// TIA Portal project "Dual_Pump_Pressure_Control" (V20)

(* hardware
DEVICE "S7-1500/ET200MP station_1"  S7-1500 station
   slot 0: "Rail_0"  Rack  6ES7 590-1***0-0AA0
   slot 1: "PLC_PumpStation"  CPU 1511-1 PN  6ES7 511-1AL03-0AB0  V4.0
      slot 3: "CPU display_1"  6ES7591-1AA00-0AA0
      slot 32768: "PROFINET interface_1"  X1
         slot 32769: "Port_1"  X1 P1
         slot 32770: "Port_2"  X1 P2
      slot 34817: "Virtual CP interface port_1"  Virtual CP interface port  Virtual CP interface port FW V4.0
DEVICE "HMI_PumpStation"  TP1500 Comfort
   slot 0: "HMI_PumpStation"  TP1500 Comfort  6AV2 124-0QC02-0AX0  17.0.0.0
   slot 1: "HMI_RT_1"  TP1500 Comfort  6AV2 124-0QC02-0AX0  17.0.0.0
   slot 5: "HMI_PumpStation.IE_CP_1"  PROFINET Interface  17.0.0.0
      slot 1: "PROFINET Interface_1"  PROFINET Interface
         slot 1: "Port_1"  Port
         slot 2: "Port_2"  Port
   slot 6: "HMI_PumpStation.IE_CP_2"  PROFINET Interface  17.0.0.0
      slot 1: "PROFINET Interface_GBit"  PROFINET Interface
         slot 1: "Port_1"  Port
   slot 7: "HMI_PumpStation.MPI/DP_CP_1"  MPI/DP Interface  17.0.0.0
DEVICE "SCADA_PumpStation"  SIMATIC PC station
   slot 0: "SIMATIC PC station"  Rail  SIMATIC PC-Station  V1.0
      slot 125: "Stationmanager"  Station_Manager  V6.0.4
   slot 1: "HMI_RT_2"  WinCC Unified PC RT  6AV2 155-xxxxx-xxxx  20.0.0.0
   slot 2: "IE general_1"  IE General  IE_CP  V8.2.0
      slot 1: "PROFINET interface"  IEGeneral.Interface.8.2.0
*)

// ===== PLC "PLC_PumpStation"  CPU 1511-1 PN =====

DATA_BLOCK "DB_Sim"   // DB1
{ S7_Optimized_Access := 'TRUE' }
VERSION : 0.1
   VAR
      Water_Level_OK : Bool := true;
      P1_InjectFault : Bool;
      P2_InjectFault : Bool;
   END_VAR
BEGIN
END_DATA_BLOCK

DATA_BLOCK "DB_IO"   // DB2
{ S7_Optimized_Access := 'TRUE' }
VERSION : 0.1
   VAR
      P1_RunCmd : Bool;
      P1_Speed_SP : Real := 0.0;
      P1_Ready : Bool;
      P1_RunningFB : Bool;
      P1_StoppedFB : Bool;
      P1_Fault : Bool;
      P2_RunCmd : Bool;
      P2_Speed_SP : Real;
      P2_Ready : Bool;
      P2_RunningFB : Bool;
      P2_StoppedFB : Bool;
      P2_Fault : Bool;
      P1_Status : Int;
      P2_Status : Int;
      AnyPumpRunning : Bool;
      Pressure_PV : Real;
      PID_Output : Real;
      PID_Enable : Bool;
      PID_Reset : Bool;
      PID_Mode : Int := 3;
   END_VAR
BEGIN
END_DATA_BLOCK

DATA_BLOCK "DB_VFD_Sim_P1"   // DB3
{ S7_Optimized_Access := 'TRUE' }
VERSION : 0.1
// stored: InstanceOfName FB_VFD_Sim
"FB_VFD_Sim"
BEGIN
END_DATA_BLOCK

DATA_BLOCK "DB_VFD_Sim_P2"   // DB4
{ S7_Optimized_Access := 'TRUE' }
VERSION : 0.1
// stored: InstanceOfName FB_VFD_Sim
"FB_VFD_Sim"
BEGIN
END_DATA_BLOCK

DATA_BLOCK "DB_HMI"   // DB5
{ S7_Optimized_Access := 'TRUE' }
VERSION : 0.1
   VAR
      Cmd_AutoMode : Bool;
      Cmd_Start : Bool;
      Cmd_Stop : Bool;
      Cmd_ManualPump : USInt := 1;
      Cmd_ManualSpeed_SP : Real := 50.0;
      Cmd_SystemReset : Bool;
      Pressure_SP : Real := 6.0;
   END_VAR
BEGIN
END_DATA_BLOCK

DATA_BLOCK "DB_PumpStation"   // DB6
{ S7_Optimized_Access := 'TRUE' }
VERSION : 0.1
// stored: InstanceOfName FB_PumpStation
"FB_PumpStation"
BEGIN
END_DATA_BLOCK

DATA_BLOCK "DB_Process_Sim"   // DB7
{ S7_Optimized_Access := 'TRUE' }
VERSION : 0.1
// stored: InstanceOfName FB_Process_Sim
"FB_Process_Sim"
BEGIN
END_DATA_BLOCK

DATA_BLOCK "DB_Alarms"   // DB9
{ S7_Optimized_Access := 'TRUE' }
VERSION : 0.1
   VAR
      AlarmWord : Word;
   END_VAR
BEGIN
END_DATA_BLOCK

FUNCTION_BLOCK "FB_VFD_Sim"   // FB1, LAD
{ S7_Optimized_Access := 'TRUE' }
VERSION : 0.1
   VAR_INPUT
      RunCmd : Bool;
      Speed_SP : Real;
      InjectFault : Bool;
   END_VAR
   VAR_OUTPUT
      Ready : Bool;
      RunningFB : Bool;
      StoppedFB : Bool;
      Fault : Bool;
      Status : Int;
   END_VAR
BEGIN

REGION Network 1: VFD Status Simulation
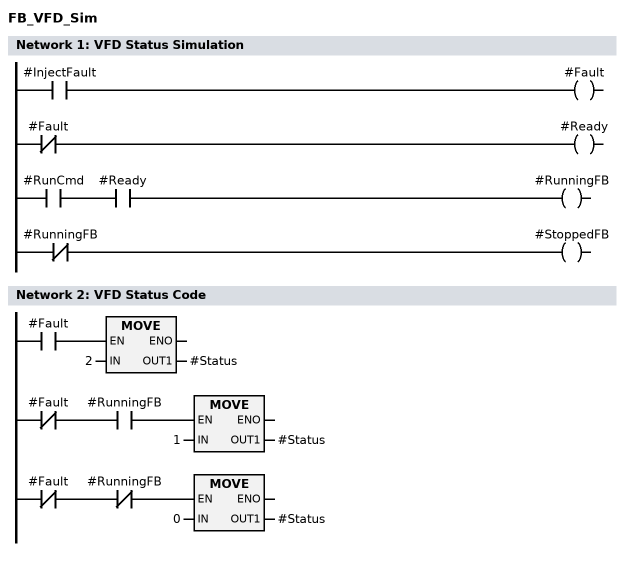
   RUNG wire#powerrail
      Contact( #InjectFault )
      Coil( #Fault )
   END_RUNG
   RUNG wire#powerrail
      I_Contact( #Fault )
      Coil( #Ready )
   END_RUNG
   RUNG wire#powerrail
      Contact( #RunCmd )
      Contact( #Ready )
      Coil( #RunningFB )
   END_RUNG
   RUNG wire#powerrail
      I_Contact( #RunningFB )
      Coil( #StoppedFB )
   END_RUNG
   // the same network as SCL:
   #Fault := #InjectFault;
   #Ready := NOT #Fault;
   #RunningFB := #RunCmd AND #Ready;
   #StoppedFB := NOT #RunningFB;
END_REGION

REGION Network 2: VFD Status Code
   RUNG wire#powerrail
      Contact( #Fault )
      Move(in := 2, out1 => #Status)
   END_RUNG
   RUNG wire#powerrail
      I_Contact( #Fault )
      Contact( #RunningFB )
      Move(in := 1, out1 => #Status)
   END_RUNG
   RUNG wire#powerrail
      I_Contact( #Fault )
      I_Contact( #RunningFB )
      Move(in := 0, out1 => #Status)
   END_RUNG
   // the same network as SCL:
   IF #Fault THEN #Status := 2; END_IF;
   IF NOT #Fault AND #RunningFB THEN #Status := 1; END_IF;
   IF NOT #Fault AND NOT #RunningFB THEN #Status := 0; END_IF;
END_REGION
END_FUNCTION_BLOCK

FUNCTION_BLOCK "FB_PumpStation"   // FB2, LAD
{ S7_Optimized_Access := 'TRUE' }
VERSION : 0.1
   VAR_INPUT
      AutoMode : Bool;
      StartCmd : Bool;
      StopCmd : Bool;
      ManualPump : USInt;
      ManualSpeed_SP : Real;
      Water_Level_OK : Bool;
      P1_Ready : Bool;
      P1_RunningFB : Bool;
      P1_StoppedFB : Bool;
      P1_Fault : Bool;
      P2_Ready : Bool;
      P2_RunningFB : Bool;
      P2_StoppedFB : Bool;
      P2_Fault : Bool;
      ResetCmd : Bool;
      AutoSpeed_SP : Real;
      Pressure_PV : Real;
   END_VAR
   VAR_OUTPUT
      P1_RunCmd : Bool;
      P1_Speed_SP : Real;
      P2_RunCmd : Bool;
      P2_Speed_SP : Real;
      HighPressureWarning : Bool;
   END_VAR
   VAR
      State : Int;
      ActivePump : USInt;
      AutoModePrevious : Bool;
      NextDutyPump : USInt := 1;
      FailoverUsed : Bool;
      StartEdge : R_TRIG;
   END_VAR
   VAR_TEMP
      ModeChanged : Bool;
      StartPulse : Bool;
      ManualStartAllowed : Bool;
      P1_StartAllowed : Bool;
      P2_StartAllowed : Bool;
      AutoStartAllowed : Bool;
      AutoP1_Available : Bool;
      AutoP2_Available : Bool;
      SpeedCommand : Real;
   END_VAR
   VAR_TEMP   // added for the SCL form of the ladder/FBD networks
      _w1 : Bool;
      _w2 : Bool;
      _w3 : Bool;
   END_VAR
BEGIN

REGION Network 1: Operating Mode Change Detection
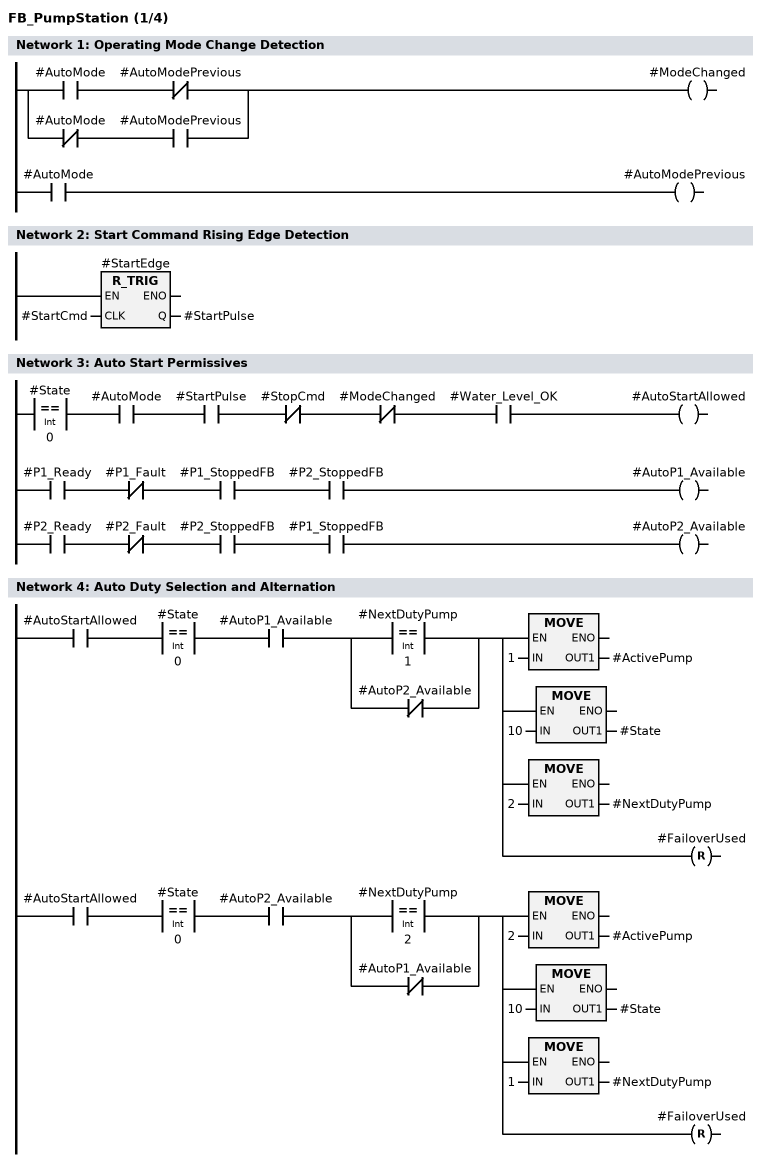
   RUNG wire#powerrail
      Contact( #AutoMode )
      I_Contact( #AutoModePrevious )
      wire#w1
      Coil( #ModeChanged )
   END_RUNG
   RUNG wire#powerrail
      I_Contact( #AutoMode )
      Contact( #AutoModePrevious )
   END_RUNG wire#w1
   RUNG wire#powerrail
      Contact( #AutoMode )
      Coil( #AutoModePrevious )
   END_RUNG
   // the same network as SCL:
   #ModeChanged := (#AutoMode AND NOT #AutoModePrevious) OR (NOT #AutoMode AND #AutoModePrevious);
   #AutoModePrevious := #AutoMode;
END_REGION

REGION Network 2: Start Command Rising Edge Detection
   #StartEdge(CLK := #StartCmd, Q => #StartPulse);   // R_TRIG
END_REGION

REGION Network 3: Auto Start Permissives
   RUNG wire#powerrail
      { S7_Templates := "SrcType := Int" } EQ_Contact(in1 := #State, in2 := 0)
      Contact( #AutoMode )
      Contact( #StartPulse )
      I_Contact( #StopCmd )
      I_Contact( #ModeChanged )
      Contact( #Water_Level_OK )
      Coil( #AutoStartAllowed )
   END_RUNG
   RUNG wire#powerrail
      Contact( #P1_Ready )
      I_Contact( #P1_Fault )
      Contact( #P1_StoppedFB )
      Contact( #P2_StoppedFB )
      Coil( #AutoP1_Available )
   END_RUNG
   RUNG wire#powerrail
      Contact( #P2_Ready )
      I_Contact( #P2_Fault )
      Contact( #P2_StoppedFB )
      Contact( #P1_StoppedFB )
      Coil( #AutoP2_Available )
   END_RUNG
   // the same network as SCL:
   #AutoStartAllowed := (#State = 0) AND #AutoMode AND #StartPulse AND NOT #StopCmd AND NOT #ModeChanged AND #Water_Level_OK;
   #AutoP1_Available := #P1_Ready AND NOT #P1_Fault AND #P1_StoppedFB AND #P2_StoppedFB;
   #AutoP2_Available := #P2_Ready AND NOT #P2_Fault AND #P2_StoppedFB AND #P1_StoppedFB;
END_REGION

REGION Network 4: Auto Duty Selection and Alternation
   RUNG wire#powerrail
      Contact( #AutoStartAllowed )
      { S7_Templates := "SrcType := Int" } EQ_Contact(in1 := #State, in2 := 0)
      Contact( #AutoP1_Available )
      wire#w1
      { S7_Templates := "SrcType := Int" } EQ_Contact(in1 := #NextDutyPump, in2 := 1)
      wire#w2
      Move(in := 1, out1 => #ActivePump)
   END_RUNG
   RUNG wire#w1
      I_Contact( #AutoP2_Available )
   END_RUNG wire#w2
   RUNG wire#w2
      Move(in := 10, out1 => #State)
   END_RUNG
   RUNG wire#w2
      Move(in := 2, out1 => #NextDutyPump)
   END_RUNG
   RUNG wire#w2
      R_Coil( #FailoverUsed )
   END_RUNG
   RUNG wire#powerrail
      Contact( #AutoStartAllowed )
      { S7_Templates := "SrcType := Int" } EQ_Contact(in1 := #State, in2 := 0)
      Contact( #AutoP2_Available )
      wire#w3
      { S7_Templates := "SrcType := Int" } EQ_Contact(in1 := #NextDutyPump, in2 := 2)
      wire#w4
      Move(in := 2, out1 => #ActivePump)
   END_RUNG
   RUNG wire#w3
      I_Contact( #AutoP1_Available )
   END_RUNG wire#w4
   RUNG wire#w4
      Move(in := 10, out1 => #State)
   END_RUNG
   RUNG wire#w4
      Move(in := 1, out1 => #NextDutyPump)
   END_RUNG
   RUNG wire#w4
      R_Coil( #FailoverUsed )
   END_RUNG
   // the same network as SCL:
   IF #AutoStartAllowed AND (#State = 0) AND #AutoP1_Available AND ((#NextDutyPump = 1) OR NOT #AutoP2_Available) THEN
       #ActivePump := 1;
   END_IF;
   #_w1 := #AutoStartAllowed AND (#State = 0) AND #AutoP1_Available AND ((#NextDutyPump = 1) OR NOT #AutoP2_Available);
   IF #_w1 THEN
       #State := 10;
       #NextDutyPump := 2;
       #FailoverUsed := FALSE;
   END_IF;
   IF #AutoStartAllowed AND (#State = 0) AND #AutoP2_Available AND ((#NextDutyPump = 2) OR NOT #AutoP1_Available) THEN
       #ActivePump := 2;
   END_IF;
   #_w2 := #AutoStartAllowed AND (#State = 0) AND #AutoP2_Available AND ((#NextDutyPump = 2) OR NOT #AutoP1_Available);
   IF #_w2 THEN
       #State := 10;
       #NextDutyPump := 1;
       #FailoverUsed := FALSE;
   END_IF;
END_REGION

REGION Network 5: Manual Start Permissives
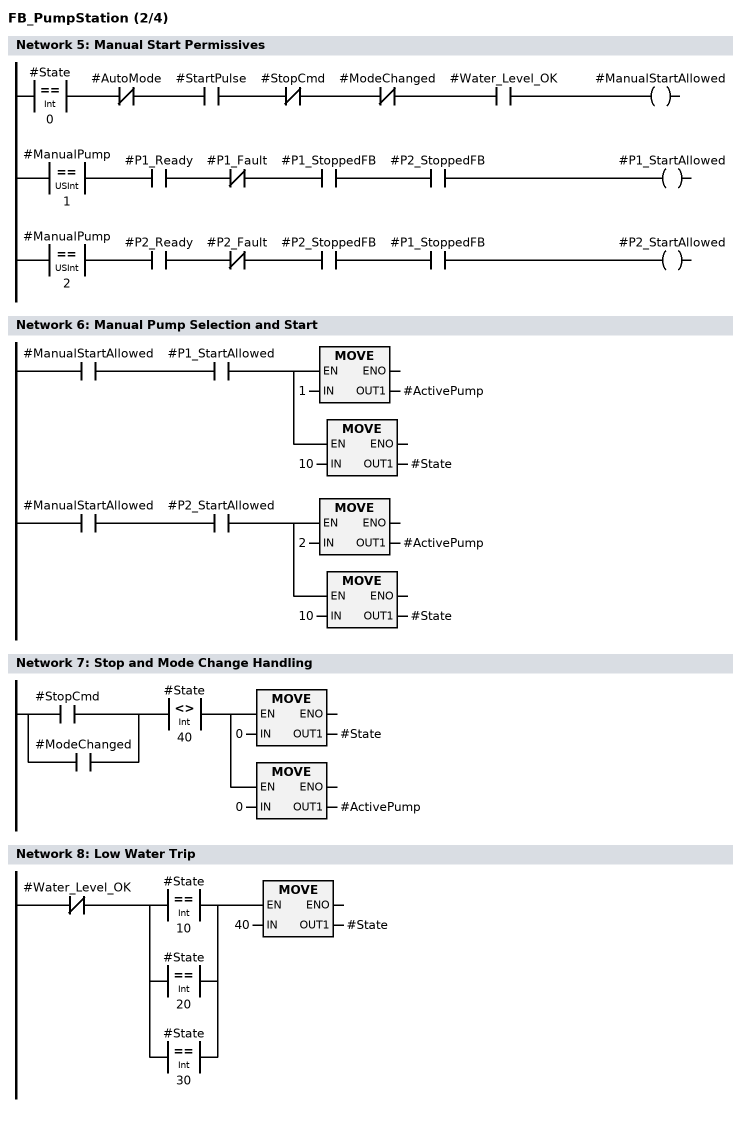
   RUNG wire#powerrail
      { S7_Templates := "SrcType := Int" } EQ_Contact(in1 := #State, in2 := 0)
      I_Contact( #AutoMode )
      Contact( #StartPulse )
      I_Contact( #StopCmd )
      I_Contact( #ModeChanged )
      Contact( #Water_Level_OK )
      Coil( #ManualStartAllowed )
   END_RUNG
   RUNG wire#powerrail
      { S7_Templates := "SrcType := USInt" } EQ_Contact(in1 := #ManualPump, in2 := 1)
      Contact( #P1_Ready )
      I_Contact( #P1_Fault )
      Contact( #P1_StoppedFB )
      Contact( #P2_StoppedFB )
      Coil( #P1_StartAllowed )
   END_RUNG
   RUNG wire#powerrail
      { S7_Templates := "SrcType := USInt" } EQ_Contact(in1 := #ManualPump, in2 := 2)
      Contact( #P2_Ready )
      I_Contact( #P2_Fault )
      Contact( #P2_StoppedFB )
      Contact( #P1_StoppedFB )
      Coil( #P2_StartAllowed )
   END_RUNG
   // the same network as SCL:
   #ManualStartAllowed := (#State = 0) AND NOT #AutoMode AND #StartPulse AND NOT #StopCmd AND NOT #ModeChanged AND #Water_Level_OK;
   #P1_StartAllowed := (#ManualPump = 1) AND #P1_Ready AND NOT #P1_Fault AND #P1_StoppedFB AND #P2_StoppedFB;
   #P2_StartAllowed := (#ManualPump = 2) AND #P2_Ready AND NOT #P2_Fault AND #P2_StoppedFB AND #P1_StoppedFB;
END_REGION

REGION Network 6: Manual Pump Selection and Start
   RUNG wire#powerrail
      Contact( #ManualStartAllowed )
      Contact( #P1_StartAllowed )
      wire#w1
      Move(in := 1, out1 => #ActivePump)
   END_RUNG
   RUNG wire#w1
      Move(in := 10, out1 => #State)
   END_RUNG
   RUNG wire#powerrail
      Contact( #ManualStartAllowed )
      Contact( #P2_StartAllowed )
      wire#w2
      Move(in := 2, out1 => #ActivePump)
   END_RUNG
   RUNG wire#w2
      Move(in := 10, out1 => #State)
   END_RUNG
   // the same network as SCL:
   IF #ManualStartAllowed AND #P1_StartAllowed THEN
       #ActivePump := 1;
       #State := 10;
   END_IF;
   IF #ManualStartAllowed AND #P2_StartAllowed THEN
       #ActivePump := 2;
       #State := 10;
   END_IF;
END_REGION

REGION Network 7: Stop and Mode Change Handling
   RUNG wire#powerrail
      Contact( #StopCmd )
      wire#w1
      { S7_Templates := "SrcType := Int" } NE_Contact(in1 := #State, in2 := 40)
      wire#w2
      Move(in := 0, out1 => #State)
   END_RUNG
   RUNG wire#powerrail
      Contact( #ModeChanged )
   END_RUNG wire#w1
   RUNG wire#w2
      Move(in := 0, out1 => #ActivePump)
   END_RUNG
   // the same network as SCL:
   #_w1 := (#StopCmd OR #ModeChanged) AND (#State <> 40);
   IF #_w1 THEN
       #State := 0;
       #ActivePump := 0;
   END_IF;
END_REGION

REGION Network 8: Low Water Trip
   RUNG wire#powerrail
      I_Contact( #Water_Level_OK )
      wire#w1
      { S7_Templates := "SrcType := Int" } EQ_Contact(in1 := #State, in2 := 10)
      wire#w2
      Move(in := 40, out1 => #State)
   END_RUNG
   RUNG wire#w1
      { S7_Templates := "SrcType := Int" } EQ_Contact(in1 := #State, in2 := 20)
   END_RUNG wire#w2
   RUNG wire#w1
      { S7_Templates := "SrcType := Int" } EQ_Contact(in1 := #State, in2 := 30)
   END_RUNG wire#w2
   // the same network as SCL:
   IF NOT #Water_Level_OK AND ((#State = 10) OR (#State = 20) OR (#State = 30)) THEN #State := 40; END_IF;
END_REGION

REGION Network 9: High Pressure Warning and Trip
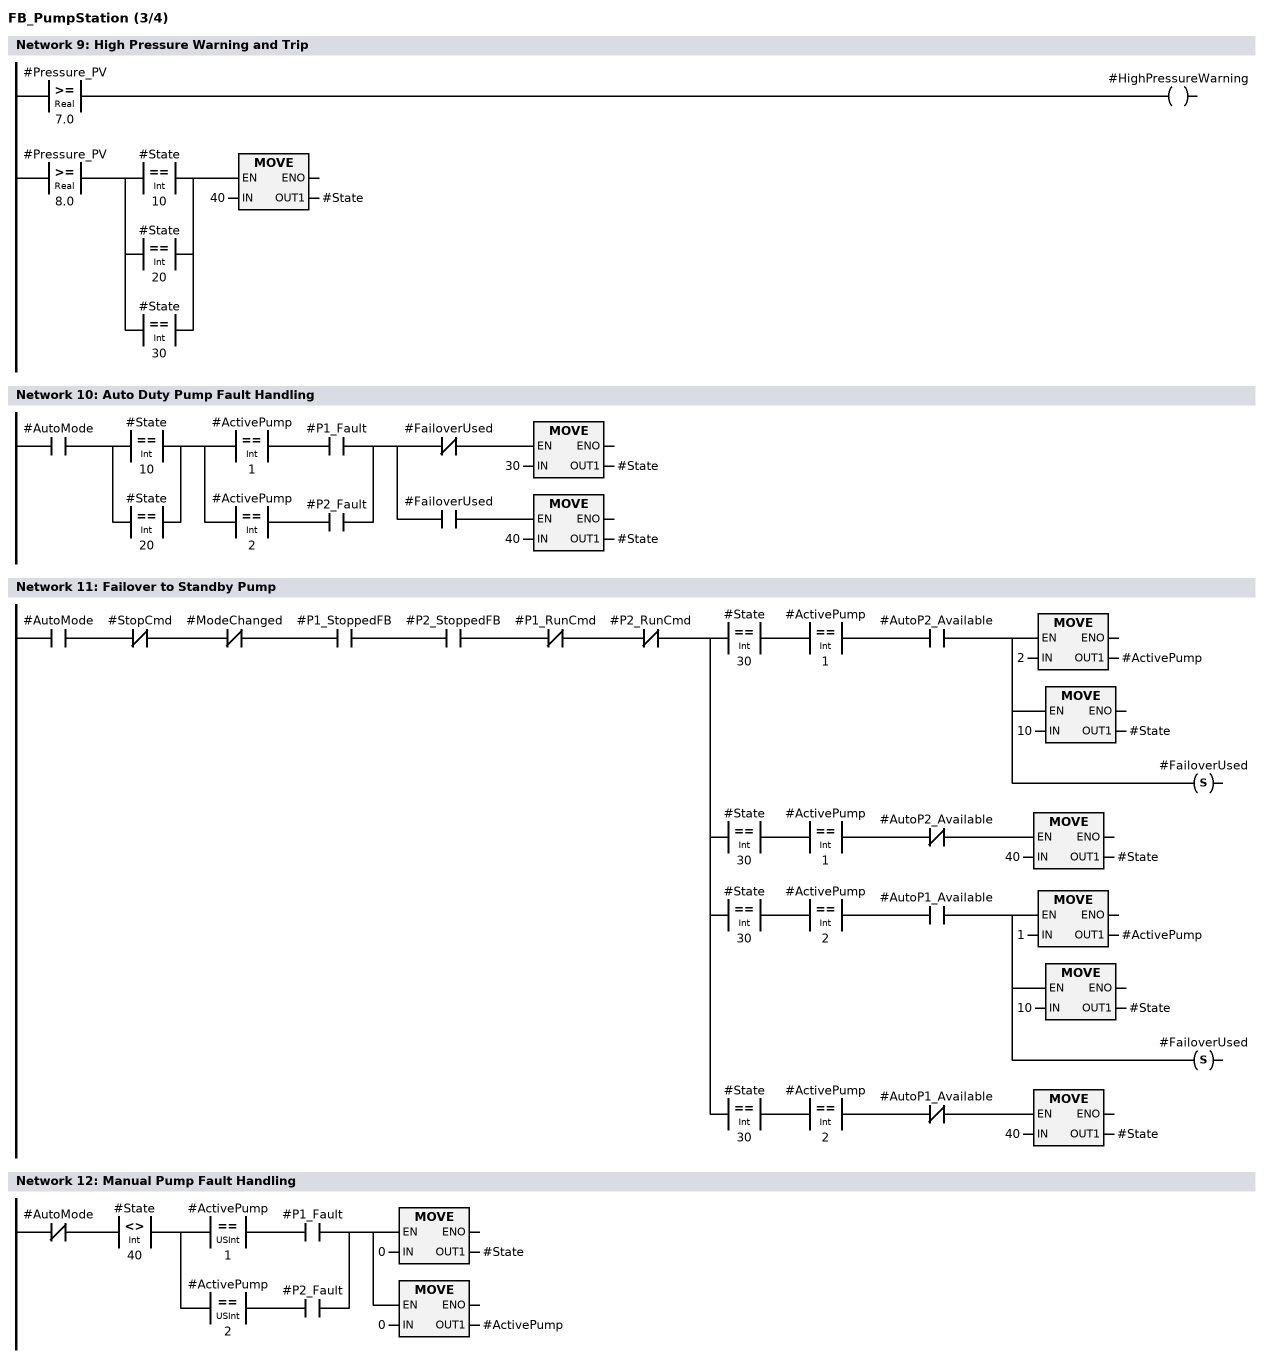
   RUNG wire#powerrail
      { S7_Templates := "SrcType := Real" } GE_Contact(in1 := #Pressure_PV, in2 := 7.0)
      Coil( #HighPressureWarning )
   END_RUNG
   RUNG wire#powerrail
      { S7_Templates := "SrcType := Real" } GE_Contact(in1 := #Pressure_PV, in2 := 8.0)
      wire#w1
      { S7_Templates := "SrcType := Int" } EQ_Contact(in1 := #State, in2 := 10)
      wire#w2
      Move(in := 40, out1 => #State)
   END_RUNG
   RUNG wire#w1
      { S7_Templates := "SrcType := Int" } EQ_Contact(in1 := #State, in2 := 20)
   END_RUNG wire#w2
   RUNG wire#w1
      { S7_Templates := "SrcType := Int" } EQ_Contact(in1 := #State, in2 := 30)
   END_RUNG wire#w2
   // the same network as SCL:
   #HighPressureWarning := #Pressure_PV >= 7.0;
   IF (#Pressure_PV >= 8.0) AND ((#State = 10) OR (#State = 20) OR (#State = 30)) THEN #State := 40; END_IF;
END_REGION

REGION Network 10: Auto Duty Pump Fault Handling
   RUNG wire#powerrail
      Contact( #AutoMode )
      wire#w1
      { S7_Templates := "SrcType := Int" } EQ_Contact(in1 := #State, in2 := 10)
      wire#w2
      { S7_Templates := "SrcType := Int" } EQ_Contact(in1 := #ActivePump, in2 := 1)
      Contact( #P1_Fault )
      wire#w3
      I_Contact( #FailoverUsed )
      Move(in := 30, out1 => #State)
   END_RUNG
   RUNG wire#w1
      { S7_Templates := "SrcType := Int" } EQ_Contact(in1 := #State, in2 := 20)
   END_RUNG wire#w2
   RUNG wire#w2
      { S7_Templates := "SrcType := Int" } EQ_Contact(in1 := #ActivePump, in2 := 2)
      Contact( #P2_Fault )
   END_RUNG wire#w3
   RUNG wire#w3
      Contact( #FailoverUsed )
      Move(in := 40, out1 => #State)
   END_RUNG
   // the same network as SCL:
   #_w1 := #AutoMode AND ((#State = 10) OR (#State = 20)) AND (((#ActivePump = 1) AND #P1_Fault) OR ((#ActivePump = 2) AND #P2_Fault));
   IF #_w1 AND NOT #FailoverUsed THEN #State := 30; END_IF;
   IF #_w1 AND #FailoverUsed THEN #State := 40; END_IF;
END_REGION

REGION Network 11: Failover to Standby Pump
   RUNG wire#powerrail
      Contact( #AutoMode )
      I_Contact( #StopCmd )
      I_Contact( #ModeChanged )
      Contact( #P1_StoppedFB )
      Contact( #P2_StoppedFB )
      I_Contact( #P1_RunCmd )
      I_Contact( #P2_RunCmd )
      wire#w1
      { S7_Templates := "SrcType := Int" } EQ_Contact(in1 := #State, in2 := 30)
      { S7_Templates := "SrcType := Int" } EQ_Contact(in1 := #ActivePump, in2 := 1)
      Contact( #AutoP2_Available )
      wire#w2
      Move(in := 2, out1 => #ActivePump)
   END_RUNG
   RUNG wire#w2
      Move(in := 10, out1 => #State)
   END_RUNG
   RUNG wire#w2
      S_Coil( #FailoverUsed )
   END_RUNG
   RUNG wire#w1
      { S7_Templates := "SrcType := Int" } EQ_Contact(in1 := #State, in2 := 30)
      { S7_Templates := "SrcType := Int" } EQ_Contact(in1 := #ActivePump, in2 := 1)
      I_Contact( #AutoP2_Available )
      Move(in := 40, out1 => #State)
   END_RUNG
   RUNG wire#w1
      { S7_Templates := "SrcType := Int" } EQ_Contact(in1 := #State, in2 := 30)
      { S7_Templates := "SrcType := Int" } EQ_Contact(in1 := #ActivePump, in2 := 2)
      Contact( #AutoP1_Available )
      wire#w3
      Move(in := 1, out1 => #ActivePump)
   END_RUNG
   RUNG wire#w3
      Move(in := 10, out1 => #State)
   END_RUNG
   RUNG wire#w3
      S_Coil( #FailoverUsed )
   END_RUNG
   RUNG wire#w1
      { S7_Templates := "SrcType := Int" } EQ_Contact(in1 := #State, in2 := 30)
      { S7_Templates := "SrcType := Int" } EQ_Contact(in1 := #ActivePump, in2 := 2)
      I_Contact( #AutoP1_Available )
      Move(in := 40, out1 => #State)
   END_RUNG
   // the same network as SCL:
   #_w1 := #AutoMode AND NOT #StopCmd AND NOT #ModeChanged AND #P1_StoppedFB AND #P2_StoppedFB AND NOT #P1_RunCmd AND NOT #P2_RunCmd;
   #_w2 := #_w1 AND (#State = 30) AND (#ActivePump = 1) AND #AutoP2_Available;
   IF #_w2 THEN
       #ActivePump := 2;
       #State := 10;
       #FailoverUsed := TRUE;
   END_IF;
   IF #_w1 AND (#State = 30) AND (#ActivePump = 1) AND NOT #AutoP2_Available THEN #State := 40; END_IF;
   #_w3 := #_w1 AND (#State = 30) AND (#ActivePump = 2) AND #AutoP1_Available;
   IF #_w3 THEN
       #ActivePump := 1;
       #State := 10;
       #FailoverUsed := TRUE;
   END_IF;
   IF #_w1 AND (#State = 30) AND (#ActivePump = 2) AND NOT #AutoP1_Available THEN #State := 40; END_IF;
END_REGION

REGION Network 12: Manual Pump Fault Handling
   RUNG wire#powerrail
      I_Contact( #AutoMode )
      { S7_Templates := "SrcType := Int" } NE_Contact(in1 := #State, in2 := 40)
      wire#w1
      { S7_Templates := "SrcType := USInt" } EQ_Contact(in1 := #ActivePump, in2 := 1)
      Contact( #P1_Fault )
      wire#w2
      Move(in := 0, out1 => #State)
   END_RUNG
   RUNG wire#w1
      { S7_Templates := "SrcType := USInt" } EQ_Contact(in1 := #ActivePump, in2 := 2)
      Contact( #P2_Fault )
   END_RUNG wire#w2
   RUNG wire#w2
      Move(in := 0, out1 => #ActivePump)
   END_RUNG
   // the same network as SCL:
   #_w1 := NOT #AutoMode AND (#State <> 40) AND (((#ActivePump = 1) AND #P1_Fault) OR ((#ActivePump = 2) AND #P2_Fault));
   IF #_w1 THEN
       #State := 0;
       #ActivePump := 0;
   END_IF;
END_REGION

REGION Network 13: System Trip Reset
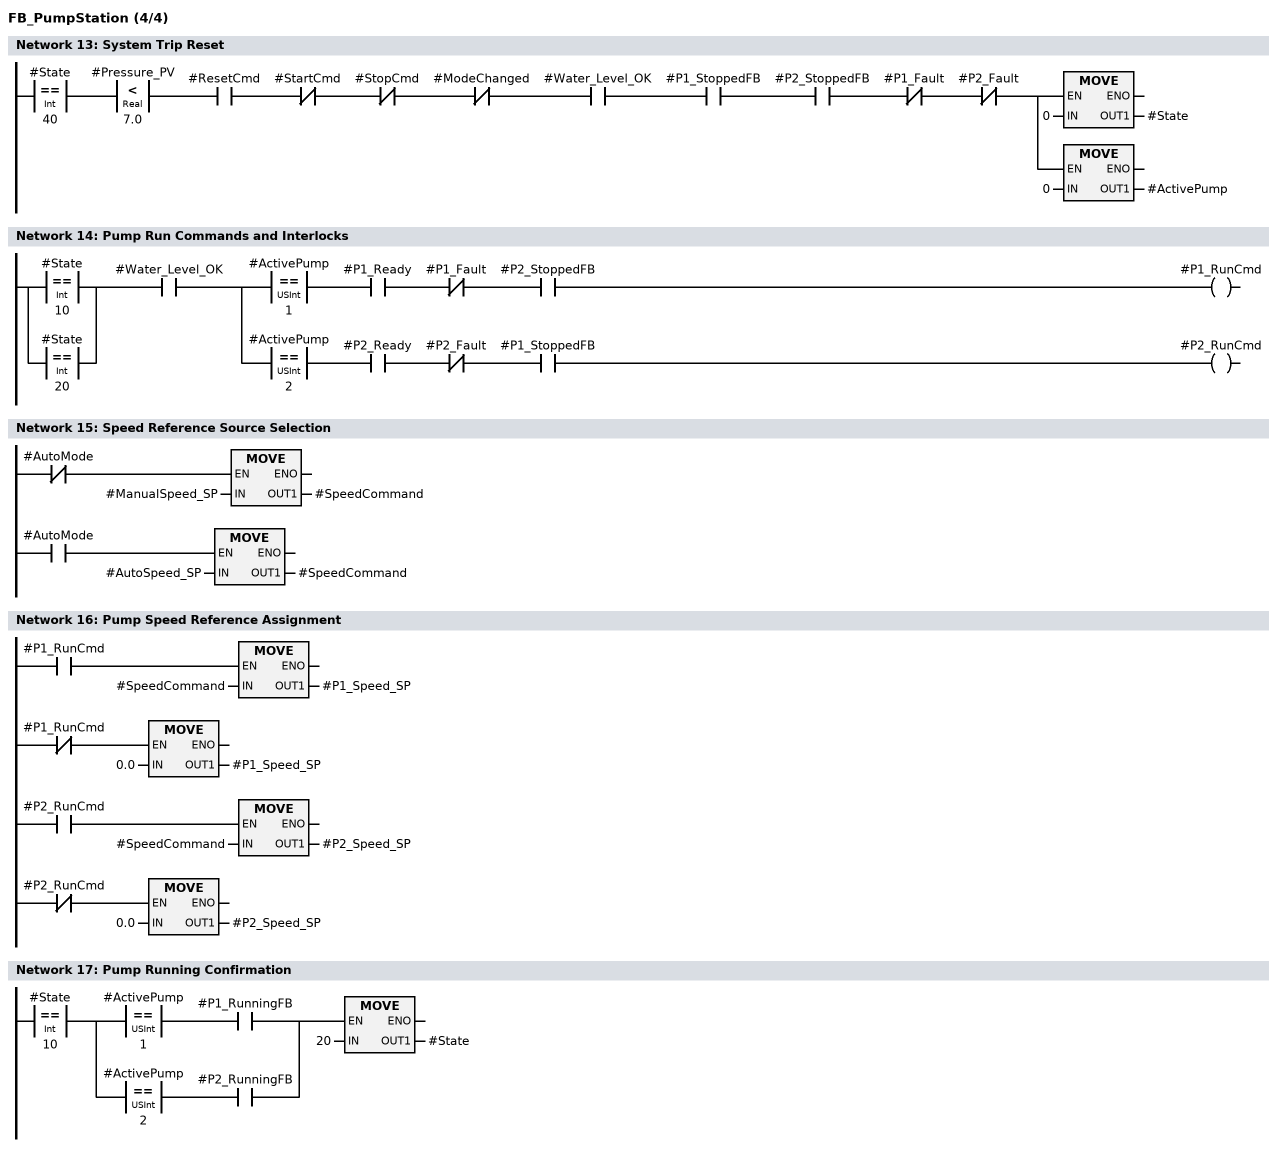
   RUNG wire#powerrail
      { S7_Templates := "SrcType := Int" } EQ_Contact(in1 := #State, in2 := 40)
      { S7_Templates := "SrcType := Real" } LT_Contact(in1 := #Pressure_PV, in2 := 7.0)
      Contact( #ResetCmd )
      I_Contact( #StartCmd )
      I_Contact( #StopCmd )
      I_Contact( #ModeChanged )
      Contact( #Water_Level_OK )
      Contact( #P1_StoppedFB )
      Contact( #P2_StoppedFB )
      I_Contact( #P1_Fault )
      I_Contact( #P2_Fault )
      wire#w1
      Move(in := 0, out1 => #State)
   END_RUNG
   RUNG wire#w1
      Move(in := 0, out1 => #ActivePump)
   END_RUNG
   // the same network as SCL:
   #_w1 := (#State = 40) AND (#Pressure_PV < 7.0) AND #ResetCmd AND NOT #StartCmd AND NOT #StopCmd AND NOT #ModeChanged AND #Water_Level_OK AND #P1_StoppedFB AND #P2_StoppedFB AND NOT #P1_Fault AND NOT #P2_Fault;
   IF #_w1 THEN
       #State := 0;
       #ActivePump := 0;
   END_IF;
END_REGION

REGION Network 14: Pump Run Commands and Interlocks
   RUNG wire#powerrail
      { S7_Templates := "SrcType := Int" } EQ_Contact(in1 := #State, in2 := 10)
      wire#w1
      Contact( #Water_Level_OK )
      wire#w2
      { S7_Templates := "SrcType := USInt" } EQ_Contact(in1 := #ActivePump, in2 := 1)
      Contact( #P1_Ready )
      I_Contact( #P1_Fault )
      Contact( #P2_StoppedFB )
      Coil( #P1_RunCmd )
   END_RUNG
   RUNG wire#powerrail
      { S7_Templates := "SrcType := Int" } EQ_Contact(in1 := #State, in2 := 20)
   END_RUNG wire#w1
   RUNG wire#w2
      { S7_Templates := "SrcType := USInt" } EQ_Contact(in1 := #ActivePump, in2 := 2)
      Contact( #P2_Ready )
      I_Contact( #P2_Fault )
      Contact( #P1_StoppedFB )
      Coil( #P2_RunCmd )
   END_RUNG
   // the same network as SCL:
   #_w1 := ((#State = 10) OR (#State = 20)) AND #Water_Level_OK;
   #P1_RunCmd := #_w1 AND (#ActivePump = 1) AND #P1_Ready AND NOT #P1_Fault AND #P2_StoppedFB;
   #P2_RunCmd := #_w1 AND (#ActivePump = 2) AND #P2_Ready AND NOT #P2_Fault AND #P1_StoppedFB;
END_REGION

REGION Network 15: Speed Reference Source Selection
   RUNG wire#powerrail
      I_Contact( #AutoMode )
      Move(in := #ManualSpeed_SP, out1 => #SpeedCommand)
   END_RUNG
   RUNG wire#powerrail
      Contact( #AutoMode )
      Move(in := #AutoSpeed_SP, out1 => #SpeedCommand)
   END_RUNG
   // the same network as SCL:
   IF NOT #AutoMode THEN #SpeedCommand := #ManualSpeed_SP; END_IF;
   IF #AutoMode THEN #SpeedCommand := #AutoSpeed_SP; END_IF;
END_REGION

REGION Network 16: Pump Speed Reference Assignment
   RUNG wire#powerrail
      Contact( #P1_RunCmd )
      Move(in := #SpeedCommand, out1 => #P1_Speed_SP)
   END_RUNG
   RUNG wire#powerrail
      I_Contact( #P1_RunCmd )
      Move(in := 0.0, out1 => #P1_Speed_SP)
   END_RUNG
   RUNG wire#powerrail
      Contact( #P2_RunCmd )
      Move(in := #SpeedCommand, out1 => #P2_Speed_SP)
   END_RUNG
   RUNG wire#powerrail
      I_Contact( #P2_RunCmd )
      Move(in := 0.0, out1 => #P2_Speed_SP)
   END_RUNG
   // the same network as SCL:
   IF #P1_RunCmd THEN #P1_Speed_SP := #SpeedCommand; END_IF;
   IF NOT #P1_RunCmd THEN #P1_Speed_SP := 0.0; END_IF;
   IF #P2_RunCmd THEN #P2_Speed_SP := #SpeedCommand; END_IF;
   IF NOT #P2_RunCmd THEN #P2_Speed_SP := 0.0; END_IF;
END_REGION

REGION Network 17: Pump Running Confirmation
   RUNG wire#powerrail
      { S7_Templates := "SrcType := Int" } EQ_Contact(in1 := #State, in2 := 10)
      wire#w1
      { S7_Templates := "SrcType := USInt" } EQ_Contact(in1 := #ActivePump, in2 := 1)
      Contact( #P1_RunningFB )
      wire#w2
      Move(in := 20, out1 => #State)
   END_RUNG
   RUNG wire#w1
      { S7_Templates := "SrcType := USInt" } EQ_Contact(in1 := #ActivePump, in2 := 2)
      Contact( #P2_RunningFB )
   END_RUNG wire#w2
   // the same network as SCL:
   IF (#State = 10) AND (((#ActivePump = 1) AND #P1_RunningFB) OR ((#ActivePump = 2) AND #P2_RunningFB)) THEN
       #State := 20;
   END_IF;
END_REGION
END_FUNCTION_BLOCK

FUNCTION_BLOCK "FB_Process_Sim"   // FB3, SCL
{ S7_Optimized_Access := 'TRUE' }
VERSION : 0.1
   VAR_INPUT
      P1_RunningFB : Bool;
      P1_Speed_SP : Real;
      P2_RunningFB : Bool;
      P2_Speed_SP : Real;
      CycleTime_s : Real := 0.1;
   END_VAR
   VAR_OUTPUT
      Pressure_PV : Real;
   END_VAR
   VAR_TEMP
      EffectiveSpeed : Real;
      TargetPressure : Real;
   END_VAR
BEGIN
   // 1. Get the speed setpoint of the running pump
   #EffectiveSpeed := 0.0;

   IF #P1_RunningFB THEN
       #EffectiveSpeed := #P1_Speed_SP;
   ELSIF #P2_RunningFB THEN
       #EffectiveSpeed := #P2_Speed_SP;
   END_IF;

   // 2. Limit the effective speed to 0–100%
   #EffectiveSpeed := LIMIT(
                            MN := 0.0,
                            IN := #EffectiveSpeed,
                            MX := 100.0
   );

   // 3. Calculate target pressure: 100% speed corresponds to 10 bar
   #TargetPressure := #EffectiveSpeed * 0.1;

   // 4. Simulate a first-order pressure response with a 3-second time constant
   #Pressure_PV := #Pressure_PV
   + (#TargetPressure - #Pressure_PV) * (#CycleTime_s / 3.0);

   // 5. Limit the pressure to 0–10 bar
   #Pressure_PV := LIMIT(
                         MN := 0.0,
                         IN := #Pressure_PV,
                         MX := 10.0
   );
END_FUNCTION_BLOCK

ORGANIZATION_BLOCK "Main"   // OB1, LAD, ProgramCycle
TITLE = "Main Program Sweep (Cycle)"
{ S7_Optimized_Access := 'TRUE' }
VERSION : 0.1
   VAR_INPUT
      Initial_Call : Bool;   // Initial call of this OB
      Remanence : Bool;   // =True, if remanent data are available
   END_VAR
BEGIN

REGION Network 1: VFD Simulation and Running Status
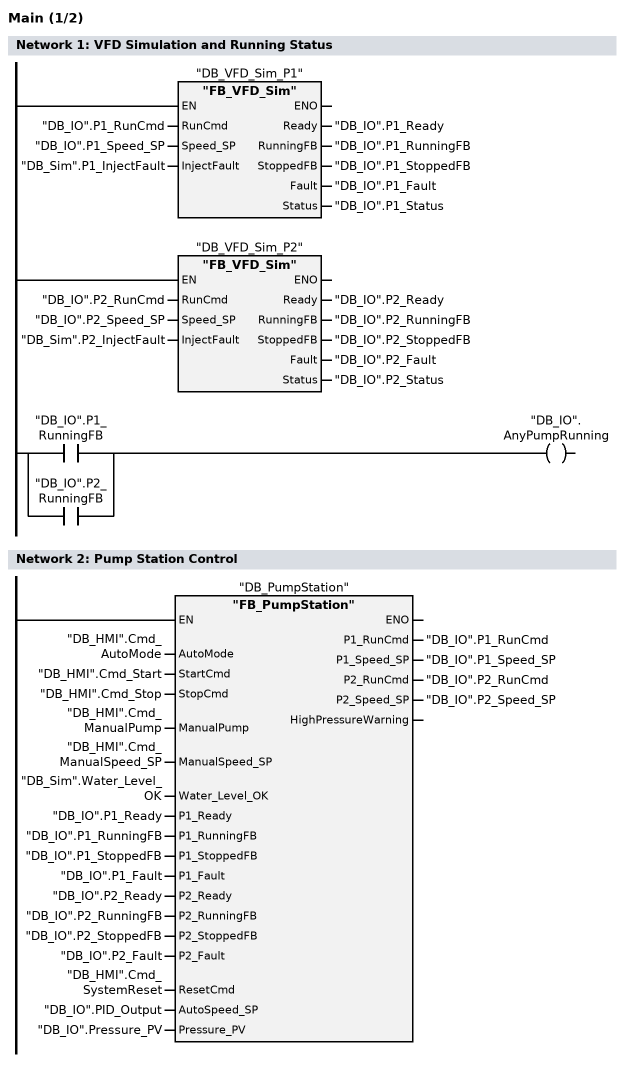
   RUNG wire#powerrail
      "DB_VFD_Sim_P1"(RunCmd := "DB_IO".P1_RunCmd, Speed_SP := "DB_IO".P1_Speed_SP, InjectFault := "DB_Sim".P1_InjectFault, Ready => "DB_IO".P1_Ready, RunningFB => "DB_IO".P1_RunningFB, StoppedFB => "DB_IO".P1_StoppedFB, Fault => "DB_IO".P1_Fault, Status => "DB_IO".P1_Status)
   END_RUNG
   RUNG wire#powerrail
      "DB_VFD_Sim_P2"(RunCmd := "DB_IO".P2_RunCmd, Speed_SP := "DB_IO".P2_Speed_SP, InjectFault := "DB_Sim".P2_InjectFault, Ready => "DB_IO".P2_Ready, RunningFB => "DB_IO".P2_RunningFB, StoppedFB => "DB_IO".P2_StoppedFB, Fault => "DB_IO".P2_Fault, Status => "DB_IO".P2_Status)
   END_RUNG
   RUNG wire#powerrail
      Contact( "DB_IO".P1_RunningFB )
      wire#w1
      Coil( "DB_IO".AnyPumpRunning )
   END_RUNG
   RUNG wire#powerrail
      Contact( "DB_IO".P2_RunningFB )
   END_RUNG wire#w1
   // the same network as SCL:
   "DB_VFD_Sim_P1"(RunCmd := "DB_IO".P1_RunCmd,   // "FB_VFD_Sim"
                   Speed_SP := "DB_IO".P1_Speed_SP,
                   InjectFault := "DB_Sim".P1_InjectFault,
                   Ready => "DB_IO".P1_Ready,
                   RunningFB => "DB_IO".P1_RunningFB,
                   StoppedFB => "DB_IO".P1_StoppedFB,
                   Fault => "DB_IO".P1_Fault,
                   Status => "DB_IO".P1_Status);
   "DB_VFD_Sim_P2"(RunCmd := "DB_IO".P2_RunCmd,   // "FB_VFD_Sim"
                   Speed_SP := "DB_IO".P2_Speed_SP,
                   InjectFault := "DB_Sim".P2_InjectFault,
                   Ready => "DB_IO".P2_Ready,
                   RunningFB => "DB_IO".P2_RunningFB,
                   StoppedFB => "DB_IO".P2_StoppedFB,
                   Fault => "DB_IO".P2_Fault,
                   Status => "DB_IO".P2_Status);
   "DB_IO".AnyPumpRunning := "DB_IO".P1_RunningFB OR "DB_IO".P2_RunningFB;
END_REGION

REGION Network 2: Pump Station Control
   RUNG wire#powerrail
      "DB_PumpStation"(AutoMode := "DB_HMI".Cmd_AutoMode, StartCmd := "DB_HMI".Cmd_Start, StopCmd := "DB_HMI".Cmd_Stop, ManualPump := "DB_HMI".Cmd_ManualPump, ManualSpeed_SP := "DB_HMI".Cmd_ManualSpeed_SP, Water_Level_OK := "DB_Sim".Water_Level_OK, P1_Ready := "DB_IO".P1_Ready, P1_RunningFB := "DB_IO".P1_RunningFB, P1_StoppedFB := "DB_IO".P1_StoppedFB, P1_Fault := "DB_IO".P1_Fault, P2_Ready := "DB_IO".P2_Ready, P2_RunningFB := "DB_IO".P2_RunningFB, P2_StoppedFB := "DB_IO".P2_StoppedFB, P2_Fault := "DB_IO".P2_Fault, ResetCmd := "DB_HMI".Cmd_SystemReset, AutoSpeed_SP := "DB_IO".PID_Output, Pressure_PV := "DB_IO".Pressure_PV, P1_RunCmd => "DB_IO".P1_RunCmd, P1_Speed_SP => "DB_IO".P1_Speed_SP, P2_RunCmd => "DB_IO".P2_RunCmd, P2_Speed_SP => "DB_IO".P2_Speed_SP, HighPressureWarning =>)
   END_RUNG
   // the same network as SCL:
   "DB_PumpStation"(AutoMode := "DB_HMI".Cmd_AutoMode,   // "FB_PumpStation"
                    StartCmd := "DB_HMI".Cmd_Start,
                    StopCmd := "DB_HMI".Cmd_Stop,
                    ManualPump := "DB_HMI".Cmd_ManualPump,
                    ManualSpeed_SP := "DB_HMI".Cmd_ManualSpeed_SP,
                    Water_Level_OK := "DB_Sim".Water_Level_OK,
                    P1_Ready := "DB_IO".P1_Ready,
                    P1_RunningFB := "DB_IO".P1_RunningFB,
                    P1_StoppedFB := "DB_IO".P1_StoppedFB,
                    P1_Fault := "DB_IO".P1_Fault,
                    P2_Ready := "DB_IO".P2_Ready,
                    P2_RunningFB := "DB_IO".P2_RunningFB,
                    P2_StoppedFB := "DB_IO".P2_StoppedFB,
                    P2_Fault := "DB_IO".P2_Fault,
                    ResetCmd := "DB_HMI".Cmd_SystemReset,
                    AutoSpeed_SP := "DB_IO".PID_Output,
                    Pressure_PV := "DB_IO".Pressure_PV,
                    P1_RunCmd => "DB_IO".P1_RunCmd,
                    P1_Speed_SP => "DB_IO".P1_Speed_SP,
                    P2_RunCmd => "DB_IO".P2_RunCmd,
                    P2_Speed_SP => "DB_IO".P2_Speed_SP);
END_REGION

REGION Network 3: HMI Alarm Mapping
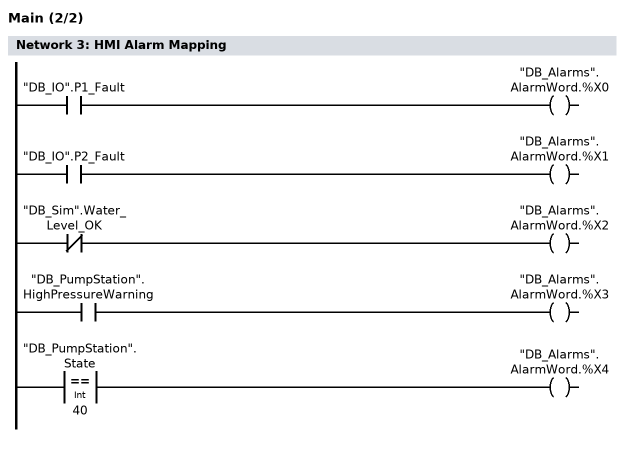
   RUNG wire#powerrail
      Contact( "DB_IO".P1_Fault )
      Coil( "DB_Alarms".AlarmWord.%X0 )
   END_RUNG
   RUNG wire#powerrail
      Contact( "DB_IO".P2_Fault )
      Coil( "DB_Alarms".AlarmWord.%X1 )
   END_RUNG
   RUNG wire#powerrail
      I_Contact( "DB_Sim".Water_Level_OK )
      Coil( "DB_Alarms".AlarmWord.%X2 )
   END_RUNG
   RUNG wire#powerrail
      Contact( "DB_PumpStation".HighPressureWarning )
      Coil( "DB_Alarms".AlarmWord.%X3 )
   END_RUNG
   RUNG wire#powerrail
      { S7_Templates := "SrcType := Int" } EQ_Contact(in1 := "DB_PumpStation".State, in2 := 40)
      Coil( "DB_Alarms".AlarmWord.%X4 )
   END_RUNG
   // the same network as SCL:
   "DB_Alarms".AlarmWord.%X0 := "DB_IO".P1_Fault;
   "DB_Alarms".AlarmWord.%X1 := "DB_IO".P2_Fault;
   "DB_Alarms".AlarmWord.%X2 := NOT "DB_Sim".Water_Level_OK;
   "DB_Alarms".AlarmWord.%X3 := "DB_PumpStation".HighPressureWarning;
   "DB_Alarms".AlarmWord.%X4 := "DB_PumpStation".State = 40;
END_REGION
END_ORGANIZATION_BLOCK

ORGANIZATION_BLOCK "OB_Process"   // OB30, LAD, CyclicInterrupt
{ S7_Optimized_Access := 'TRUE' }
VERSION : 0.1
   VAR_INPUT
      Initial_Call : Bool;   // Initial call of this OB
      Event_Count : Int;   // Events discarded
   END_VAR
BEGIN

REGION Network 1: Process Pressure Simulation
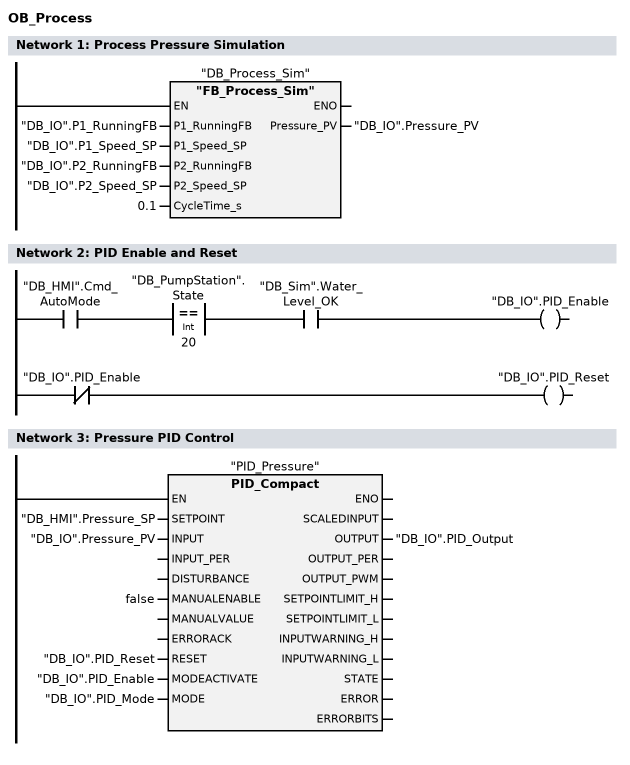
   RUNG wire#powerrail
      "DB_Process_Sim"(P1_RunningFB := "DB_IO".P1_RunningFB, P1_Speed_SP := "DB_IO".P1_Speed_SP, P2_RunningFB := "DB_IO".P2_RunningFB, P2_Speed_SP := "DB_IO".P2_Speed_SP, CycleTime_s := 0.1, Pressure_PV => "DB_IO".Pressure_PV)
   END_RUNG
   // the same network as SCL:
   "DB_Process_Sim"(P1_RunningFB := "DB_IO".P1_RunningFB,   // "FB_Process_Sim"
                    P1_Speed_SP := "DB_IO".P1_Speed_SP,
                    P2_RunningFB := "DB_IO".P2_RunningFB,
                    P2_Speed_SP := "DB_IO".P2_Speed_SP,
                    CycleTime_s := 0.1,
                    Pressure_PV => "DB_IO".Pressure_PV);
END_REGION

REGION Network 2: PID Enable and Reset
   RUNG wire#powerrail
      Contact( "DB_HMI".Cmd_AutoMode )
      { S7_Templates := "SrcType := Int" } EQ_Contact(in1 := "DB_PumpStation".State, in2 := 20)
      Contact( "DB_Sim".Water_Level_OK )
      Coil( "DB_IO".PID_Enable )
   END_RUNG
   RUNG wire#powerrail
      I_Contact( "DB_IO".PID_Enable )
      Coil( "DB_IO".PID_Reset )
   END_RUNG
   // the same network as SCL:
   "DB_IO".PID_Enable := "DB_HMI".Cmd_AutoMode AND ("DB_PumpStation".State = 20) AND "DB_Sim".Water_Level_OK;
   "DB_IO".PID_Reset := NOT "DB_IO".PID_Enable;
END_REGION

REGION Network 3: Pressure PID Control
   "PID_Pressure"(Setpoint := "DB_HMI".Pressure_SP,   // PID_Compact
                  Input := "DB_IO".Pressure_PV,
                  ManualEnable := false,
                  Reset := "DB_IO".PID_Reset,
                  ModeActivate := "DB_IO".PID_Enable,
                  Mode := "DB_IO".PID_Mode,
                  Output => "DB_IO".PID_Output);
END_REGION
END_ORGANIZATION_BLOCK

(* ===== HMI "HMI_RT_1" =====
system functions are stored by id; their names below are inferred from use
connection "HMI_Connection_3": ETHERNET, S7_1500_OMS
connection "HMI_Connection_4": ETHERNET, S7_1500_OMS

HMI tags "Default tag table"
   "DB_HMI_Cmd_ManualPump" : USInt = PLC DB_HMI.Cmd_ManualPump, 1 s
   "DB_HMI_Cmd_ManualSpeed_SP" : Real = PLC DB_HMI.Cmd_ManualSpeed_SP, 1 s
   "DB_HMI_Cmd_AutoMode" : Bool = PLC DB_HMI.Cmd_AutoMode, 1 s
   "DB_HMI_Cmd_Start" : Bool = PLC DB_HMI.Cmd_Start, 1 s
   "DB_HMI_Cmd_Stop" : Bool = PLC DB_HMI.Cmd_Stop, 1 s
   "DB_PumpStation_State" : Int = PLC DB_PumpStation.State, 1 s
   "DB_Sim_P1_InjectFault" : Bool = PLC DB_Sim.P1_InjectFault, 1 s
   "DB_Sim_P2_InjectFault" : Bool = PLC DB_Sim.P2_InjectFault, 1 s
   "DB_Sim_Water_Level_OK" : Bool = PLC DB_Sim.Water_Level_OK, 1 s
   "DB_IO_P1_Status" : Int = PLC DB_IO.P1_Status, 1 s
   "DB_IO_P2_Status" : Int = PLC DB_IO.P2_Status, 1 s
   "DB_IO_P1_RunningFB" : Bool = PLC DB_IO.P1_RunningFB, 1 s
   "DB_IO_P2_RunningFB" : Bool = PLC DB_IO.P2_RunningFB, 1 s
   "DB_IO_AnyPumpRunning" : Bool = PLC DB_IO.AnyPumpRunning, 1 s
   "DB_HMI_Cmd_SystemReset" : Bool = PLC DB_HMI.Cmd_SystemReset, 1 s
   "DB_IO_Pressure_PV" : Real = PLC DB_IO.Pressure_PV, 1 s
   "DB_HMI_Pressure_SP" : Real = PLC DB_HMI.Pressure_SP, 1 s
   "DB_Alarms_AlarmWord" : Word = PLC DB_Alarms.AlarmWord, 1 s

discrete alarms
   1: 'Lỗi VFD bơm 1', class Errors, trigger "DB_Alarms_AlarmWord" bit 0
   2: 'Lỗi VFD bơm 2', class Errors, trigger "DB_Alarms_AlarmWord" bit 1
   3: 'Mức nước không đủ', class Errors, trigger "DB_Alarms_AlarmWord" bit 2
   4: 'Cảnh báo áp suất cao ≥7 bar', class Warnings, trigger "DB_Alarms_AlarmWord" bit 3
   5: 'Hệ thống TRIPPED — cần Reset', class Errors, trigger "DB_Alarms_AlarmWord" bit 4

text list "PumpSelection": 0 'Chưa chọn'; 1 'Bơm 1'; 2 'Bơm 2'

text list "ModeSelection": 0 'Manual'; 1 'Auto'

text list "SystemState": 0 'IDLE'; 10 'STARTING'; 20 'RUNNING'; 30 'FAILOVER'; 40 'TRIPPED'

Template "Template_1" 1280x799
   Button "Template_Button" at 943,707 size 79x59; TextOff 'Text'
   Button "Template_Button_1" at 857,707 size 79x59; TextOff 'Text'
   Button "Template_Button_2" at 772,707 size 79x59; TextOff 'Text'
   Button "Template_Button_3" at 686,707 size 79x59; TextOff 'Text'
   Button "Template_Button_4" at 600,707 size 79x59; TextOff 'Text'
   Button "Template_Button_5" at 515,707 size 79x59; TextOff 'Text'
   Button "Template_Button_6" at 429,707 size 79x59; TextOff 'Text'
   Button "Template_Button_7" at 344,707 size 79x59; TextOff 'Text'
   Button "Template_Button_8" at 258,707 size 79x59; TextOff 'Text'
   Button "Template_Button_9" at 172,707 size 79x59; TextOff 'Text'
   Button "Template_Button_10" at 87,707 size 79x59; TextOff 'Text'
   Button "Template_Button_11" at 1,707 size 79x59; TextOff 'Text'

screen "Overview" 1280x799, template "Template_1"
   TextField "Text field_2" at 15,135 size 12x20; Text 'Text'
   TextField "Text field_1" at 349,11 size 631x38; Text 'Hệ thống điều khiển áp suất hai bơm'
   TextField "Text field_4" at 912,122 size 71x26; Text 'Chế độ'
   TextField "Text field_5" at 910,233 size 103x26; Text 'Chọn bơm'
   TextField "Text field_6" at 911,344 size 196x26; Text 'Tốc độ Manual (%)'
   IOField "I/O field_1" at 917,379 size 182x45; FormatPattern 999
      ProcessValue <- "DB_HMI_Cmd_ManualSpeed_SP"
   Button "Button_1" at 943,473 size 109x49; TextOff 'Start'
      on Press: SetBit("DB_HMI_Cmd_Start")
      on Release: ResetBit("DB_HMI_Cmd_Start")
   Button "Button_2" at 1091,473 size 109x49; TextOff 'Stop'
      on Press: SetBit("DB_HMI_Cmd_Stop")
      on Release: ResetBit("DB_HMI_Cmd_Stop")
   SymbolicIOField "Symbolic I/O field_3" at 714,92 size 110x19; TextOff '0'; TextOn '1'; TextList "SystemState"
      ProcessValue <- "DB_PumpStation_State"
   TextField "Text field_7" at 591,87 size 124x26; Text 'Trạng thái:'
   TextField "Text field_8" at 50,727 size 110x26; Text 'Mô phỏng'
   Switch "Switch_1" at 190,725 size 61x35; CaptionText 'Switch'; TextOff 'OFF'; TextOn 'ON'
      ProcessValue <- "DB_Sim_P1_InjectFault"
   TextField "Text field_9" at 254,730 size 103x24; Text 'Lỗi bơm 1'
   TextField "Text field_10" at 492,730 size 97x24; Text 'Lỗi bơm 2'
   Switch "Switch_2" at 419,724 size 61x35; CaptionText 'Switch'; TextOff 'OFF'; TextOn 'ON'
      ProcessValue <- "DB_Sim_P2_InjectFault"
   TextField "Text field_11" at 732,729 size 137x24; Text 'Mực nước đủ'
   Switch "Switch_3" at 665,724 size 61x35; CaptionText 'Switch'; TextOff 'OFF'; TextOn 'ON'
      ProcessValue <- "DB_Sim_Water_Level_OK"
   Rectangle "Rectangle_7" at 148,250 size 169x232
      Appearance <- "DB_Sim_Water_Level_OK"
   Rectangle "Rectangle_8" at 319,326 size 102x19
      Appearance <- "DB_IO_AnyPumpRunning"
   Rectangle "Rectangle_9" at 399,239 size 22x88
      Appearance <- "DB_IO_P1_RunningFB"
   Rectangle "Rectangle_10" at 399,344 size 22x101
      Appearance <- "DB_IO_P2_RunningFB"
   Rectangle "Rectangle_12" at 420,239 size 241x19
      Appearance <- "DB_IO_P1_RunningFB"
   TextField "Text field_14" at 198,193 size 71x23; Text 'Bồn cấp'
   Circle "Circle_1" at 483,198 size 96x96
      Appearance <- "DB_IO_P1_Status"
   TextField "Text field_12" at 499,233 size 62x23; Text 'Bơm 1'
   Rectangle "Rectangle_13" at 420,426 size 241x19
      Appearance <- "DB_IO_P2_RunningFB"
   Circle "Circle_2" at 482,382 size 96x96
      Appearance <- "DB_IO_P2_Status"
   TextField "Text field_13" at 499,418 size 62x23; Text 'Bơm 2'
   Rectangle "Rectangle_14" at 660,239 size 22x88
      Appearance <- "DB_IO_P1_RunningFB"
   Rectangle "Rectangle_15" at 660,344 size 22x101
      Appearance <- "DB_IO_P2_RunningFB"
   Rectangle "Rectangle_16" at 660,326 size 99x19
      Appearance <- "DB_IO_AnyPumpRunning"
   SymbolicIOField "Symbolic I/O field_4" at 911,159 size 189x47; TextOff '0'; TextOn '1'; TextList "ModeSelection"
      ProcessValue <- "DB_HMI_Cmd_AutoMode"
   SymbolicIOField "Symbolic I/O field_5" at 912,267 size 186x48; TextOff '0'; TextOn '1'; TextList "PumpSelection"
      ProcessValue <- "DB_HMI_Cmd_ManualPump"
   TextField "Text field_3" at 942,72 size 281x34; Text 'Điều khiển vận hành'
   Button "Button_3" at 948,545 size 251x49; TextOff 'RESET'
      on Press: SetBit("DB_HMI_Cmd_SystemReset")
      on Release: ResetBit("DB_HMI_Cmd_SystemReset")
   IOField "I/O field_2" at 147,620 size 125x68; FormatPattern 99.999
      ProcessValue <- "DB_IO_Pressure_PV"
   TextField "Text field_15" at 124,594 size 173x28; Text 'Áp suất đường ống'
   IOField "I/O field_3" at 536,616 size 125x68; FormatPattern 99.999
      ProcessValue <- "DB_HMI_Pressure_SP"
   TextField "Text field_16" at 540,592 size 79x28; Text 'Setpoint'
   TextField "Text field_17" at 244,640 size 34x28; Text 'bar'
   TextField "Text field_18" at 633,636 size 34x28; Text 'bar'
   Button "Button_4" at 26,6 size 102x44; TextOff 'Alarms'
      on Click: ActivateScreen("Alarms", 0)
   Button "Button_5" at 142,4 size 102x44; TextOff 'Trends'
      on Click: ActivateScreen("Trends", 0)

screen "Alarms" 1280x799
   AlarmView "Alarm view_1" at 50,80 size 1080x604
   Button "Button_1" at 50,16 size 109x43; TextOff 'Overview'
      on Click: ActivateScreen("Overview", 0)

screen "Trends" 1280x799
   TrendView "Trend view_1" at 39,95 size 1217x513
   Button "Button_1" at 56,18 size 159x61; TextOff 'Overview'
      on Click: ActivateScreen("Overview", 0)
*)

(* ===== HMI "HMI_RT_2" =====
connection "HMI_Connection_2": ETHERNET, ILRT_S7_1500_OMS

HMI tags "Default tag table"
   "Pressure_PV" : Real = PLC DB_IO.Pressure_PV, T1s
   "Pressure_SP" : Real = PLC DB_HMI.Pressure_SP AT %DB1.DBD0, T1s

text list "SystemTextList_ConfigErrorAlarmTextLibrary_1": 1 'NameService configuration error: Implicit deletion. Subelement instance @6%s@ must be deleted explicitly.'; 2 'NameService configuration error: Implicit deletion. Alias/Format/Unit instance @6%s@ must be deleted explicitly.'

text list "SystemTextList_ConfigErrorAlarmTextLibrary_2": 1 'EvDpManager::cleanupDeletedDatapoint - alert handler config is deleted implicitly for deleted datapoint, @3%s@'; 2 'EvDpManager::cleanupDeletedDatapoint - alert handler config is deleted implicitly but still has overrides, @3%s@'; 3 'EvDpManager::cleanupDeletedDatapoint - default value config is deleted implicitly for deleted datapoint, @3%s@'; 4 'EvDpManager::cleanupDeletedDatapoint - default value config is deleted implicitly but still has overrides, @3%s@'; 5 'EvDpManager::cleanupDeletedDatapoint - initial value config is deleted implicitly for deleted datapoint, @3%s@'; 6 'EvDpManager::cleanupDeletedDatapoint - initial value config is deleted implicitly but still has overrides, @3%s@'; 7 'EvDpManager::cleanupDeletedDatapoint - distribution config is deleted implicitly for deleted datapoint, @3%s@'; 8 'EvDpManager::cleanupDeletedDatapoint - distribution config is deleted implicitly but still has overrides, @3%s@'; 9 'EvDpManager::cleanupDeletedDatapoint - rangeCheck config is deleted implicitly for deleted datapoint, @3%s@'; 10 'EvDpManager::cleanupDeletedDatapoint - rangeCheck config is deleted implicitly but still has overrides, @3%s@'

text list "SystemTextList_ConfigErrorAlarmTextLibrary_3": 1 'The configured data point type was deleted, but a configured type is still defined for the node type: @3%s@.'; 2 'The configured data point node type was deleted in the data point type, but a configured type is still defined for the element: @3%s@.'

text list "SystemTextList_ConfigErrorAlarmTextLibrary_4": 2 'Cycles: @6%s@ does not exist'; 3 'Alarms: @6%s@ exists already'; 4 'Tags: Address @6%s@ was rejected'; 1 'Connections: @6%s@ does not exist'; 5 'Tags: Acquisition mode @6%s@ is not supported.'; 6 'Cycles: @6%s@ was deleted but associated tags exist.'; 7 'Connections: @6%s@ was deleted but associated tags exist.'; 8 'Tags: Tag @6%s@ was rejected.'; 9 'Tags: Tag @6%s@ has an invalid value.'; 0 'Connections: Connection to @6%s@ could not be established.'; 65638 'Connections: Connection to @6%s@ could not be established.'; 65639 'Connections: @6%s@ disconnected.'; 65640 'Connections: Connection to the HMI device @6%s@ is lost.'; 65641 'Connections: Connection to the PLC @6%s@ is lost.'; 65541 'Connections: Timeout while establishing the connection to @6%s@.'; 65542 'Connections: @6%s@ faulty.'; 65543 'Connections: Connection to the HMI device disconnected. Connection @5%s@ was changed.'; 65544 'Connections: Connection to the HMI device disconnected. Driver property was changed for connection @5%s@.'

text list "SystemTextList_ConfigErrorAlarmTextLibrary_5": 1 'Connections: Lifecycle monitoring cycle must be shorter than the response time.'; 2 'Connections: Cyclic services are configured but not supported by the target device.'; 3 'Connections: Change-controlled reading is configured but not supported by the target device.'; 4 'Tags: The address @6%s@ does not exist in the PLC.'; 5 'Tags: The default conversion type for the address @6%s@ could not be determined.'; 6 'Tags: Invalid conversion type'; 7 'Cycles: Invalid conversion type. Conversion is not supported at HmiCycle.'; 4096 'Connections: Version of the address @6%s@ is not supported.'; 4097 'Connections: PROFIBUS address is not supported.'; 4098 'Connections: Softbus address is not supported.'; 4099 'Connections: Address type @6%s@ is not supported.'; 4100 'Connections: Invalid connection name @6%s@. Access point is being ignored.'; 4101 'Connections: Routing is not supported. @6%s@ is not used.'; 4102 'Connections: Routing is not supported. @6%s@ is not used.'; 4103 'Connections: Invalid IP address @6%s@'; 4104 'Connections: Invalid Named Connection @6%s@. Valid format: >VMD</>connection<'; 4105 'Connections: Invalid Named Connection @6%s@. VMD connection name is too long. Only 24 characters are permitted.'; 4106 'Connections: Invalid Named Connection @6%s@. Connection name is too long. Only 32 characters are permitted.'; 4107 'Connections: Rack number @6%s@ is outside of the permitted range (0..7)'; 4108 'Connections: Invalid Named Connection @6%s@. Rack is ignored.'; 4109 'Connections: Slot number @6%s@ is outside of the permitted range (0..31)'; 4110 'Connections: Invalid Named Connection @6%s@. Slot is ignored.'; 4111 'Connection could not be established. Maximum number of available connections (@6%s@) has been exceeded.'; 4112 'Connection aborted. No sign of life in the last @4%s@ ms.'; 4113 'Connection could not be established - @4%s@'; 4114 'Connection could not be established. The address @6%s@ cannot be used.'; 4115 'Connection could not be established. Invalid address @6%s@'; 4116 'Connection could not be established - @4%s@'

text list "SystemTextList_ConfigErrorAlarmTextLibrary_6": 1 'Connection could not be established. Application instance certificate is not configured.'; 2 'Connection could not be established. Server has rejected the client certificate. OPC UA status code @4%s@.'; 3 'Connection could not be established. Internal problem in the certificate store. OPC UA status code @4%s@'; 4 'Connection could not be established. Application instance certificate could not be loaded. OPC UA status code @4%s@'; 5 'Connection could not be established. Server has not provided a certificate. @4%s@'; 6 'Connection could not be established. Validation of server certificate has failed. OPC UA status code @4%s@.'; 7 'Connection was closed. Error during alarm synchronization. OPC UA status code @4%s@.'; 8 'Connection was closed. Alarm/event subscription has failed. The number of operations on the server has been exceeded.'; 9 'Connection was closed. Alarm/event subscription has failed. The number of alarm/event subscriptions on the server has been exceeded.'; 10 'Connection could not be established. Server reports a license problem. OPC UA status code @4%s@.'; 11 'Connection could not be established. Maximum number of server sessions has been exceeded.'; 12 'Connection could not be established. Safety configuration is inconsistent. @4%s@'; 13 'Connection could not be established. The address @4%s@ cannot be used.'; 14 'Connection could not be established. OPC UA status code @4%s@'; 15 'Connection aborted. OPC UA server was stopped.'; 16 'Connection aborted. No sign of life in the last @4%s@ ms.'; 17 'Connection was closed. OPC UA server maintenance.'; 18 'Connection could not be established. Invalid configuration of the authentication mode - @4%s@'; 19 'Connection could not be established. User could not be authenticated. OPC UA status code @4%s@'; 20 'Connection could not be established. Server does not permit anonymous connection. OPC UA status code @4%s@'; 21 'Connection could not be established. Certificate problem: Error when writing the safety-relevant data to @4%s@.'; 22 'Connection could not be established. Certificate problem: Unexpected file in the folder @4%s@ cannot be removed.'; 23 'Connection could not be established. User could not be authenticated. No user or password configured.'; 24 'Connection could not be established. Unexpected length of the server certificate. @4%s@'; 25 'Connection could not be established. @4%s@ is empty.'; 26 'Connection could not be established. @4%s@ has an unexpected format.'; 27 'Connection could not be established. Server endpoints cannot be read. OPC UA status code @4%s@'; 28 'Connection could not be established. No server endpoints were found. @4%s@'; 29 'Connection could not be established. Application instance certificate could not be found.'; 30 'Connection could not be established. Unexpected format of the certificate @4%s@.'; 31 'Connection could not be established. Unexpected format of the certificate block list @4%s@.'; 32 'Connection could not be established. User could not be authenticated. An encryption detail is invalid. @4%s@'; 34 'Connection could not be established. - The configured non-transparent redundancy mode @4%s@ is not supported.'; 101 'Tags: Address @6%s@ does not exist on the server.'; 103 'Tags: Address @6%s@ cannot be accessed.'; 104 'Tags: Acquisition mode is not supported for address @6%s@.'; 201 'Alarms: Address @6%s@ does not exist on the server.'; 202 'Alarms: Address @6%s@ cannot be used. The specified range filter is not an OPC UA Event Notifier.'; 203 'Alarms: Address @6%s@ cannot be used. The specified range filter does not exist on the server.'; 204 'Alarms: Address @6%s@ cannot be used because it is not an OPC UA event type.'; 205 'Alarms: Address @6%s@ cannot be used because the OPC UA condition type is not supported.'; 206 'Alarms: Address @6%s@ cannot be used because the event type does not exist on the server.'; 207 'Alarms: Acquisition type cannot be used for address @6%s@.'; 301 'Address @6%s@ cannot be used because the version number is missing.'; 302 'Address @6%s@ cannot be used because the version number is invalid.'; 303 'Address @6%s@ cannot be used because the number of '$' delimiters is invalid.'; 304 'Address @6%s@ cannot be used because the address type is invalid.'; 305 'Unsupported version @6%s@ of the address'; 401 'Unexpected OPC UA server response: @6%s@'

text list "SystemTextList_ConfigErrorAlarmTextLibrary_7": 1 'Messages: Invalid condition string for the alarm view @6%s@.'; 2 'Messages: Invalid status tag and bit for the alarm view @6%s@.'; 3 'Messages: Invalid control tag and bit for the alarm view @6%s@.'

text list "SystemTextList_ConfigErrorAlarmTextLibrary_8": 1 'Logs: Implicit deletion. Logging tag instance @6%s@ should be deleted but there are overloaded elements.'

text list "SystemTextList_ConfigErrorAlarmTextLibrary_9": 2 'Restart of the runtime is required.'; 3 'The correct storage medium must be ejected and inserted again.'

text list "SystemTextList_ConfigErrorAlarmTextLibrary_10": 1 'CDS cache - Cache folder cannot be created or reached: @6%s@'; 2 'LOC cache - Cache folder cannot be created or reached: @6%s@'

text list "SystemTextList_ConfigErrorAlarmTextLibrary_11": 2 'and synchronization will start automatically. Shutting down either of them during synchronization will not cause data loss.'; 3 'and synchronization is scheduled for: @5%Y-%m-%d %H:%M:%S@. Shutting down either of the computers will not cause data loss.'

text list "SystemTextList_RuntimeCollaborationFailureReason_1": 0 'Unknown error (@3%s@)'; 1 'The system is not running or there is a network problem'; 2 'Runtime is not started on the target device.'; 3 'The System ID does not match the expected System ID (@3%s@)'; 4 'The Collaboration name does not match the expected Collaboration name '@3%s@''; 5 'Wrong or unknown certificate'; 6 'Revoked certificate'; 7 'The time difference is too big.'; 8 'No common supported message version'; 9 'System ID (@3%s@) already exists'; 10 'System name (@3%s@) already exists'; 11 'ID/Name in local configuration for Runtime Collaboration already exists'

text list "SystemTextList_RedundancyRecoveryFailureReason_1": 0 'Data recovery request temporarily rejected until own recovery request has been responded to.'; 1 'Data recovery request rejected. Online backup running.'; 2 'Data recovery request rejected. Connection to the Event Manager is not established.'; 3 'Data recovery request temporarily rejected until delta activation is complete.'; 4 'Data recovery request temporarily rejected until alarms and tags are retentive.'; 5 'Data recovery request rejected. The obligatory file config.level.es is missing on the computer.'; 6 'Data recovery request was canceled by the Event Manager.'; 7 'The data synchronization between the devices has failed.'

text list "SystemTextList_S7PlusAlarmTextListCollection_1": 4096 'Connections: Connection to the PLC @4%s@ is lost'; 4097 'Connections: Connection to the HMI device @4%s@ is lost'; 4098 'Connections: Maximum number of connections exceeded - @4%s@'; 4099 'Out of resources on PLC - @4%s@'; 4100 'Legitimation failed, invalid or missing password - @4%s@'; 4101 'Request to open the connection failed - @4%s@'; 4102 'Connections: Cannot connect to PLC - @4%s@'; 4103 'Request to open the connection could not be sent'; 4104 'General certificate error for PLC - @4%s@'; 4105 'PLC certificate expired for PLC - @4%s@'; 4106 'PLC certificate is revoked for PLC - @4%s@'; 4107 'PLC certificate is untrustworthy. Manual trust is possible for - @4%s@'; 4108 'PLC certificate is untrustworthy. Manual trust is not possible for - @4%s@'

text list "SystemTextList_AllenBradleyEIPAlarmTextListCollection_7": 4096 'Connection lost on PLC side - @5%s@'; 4097 'Connection lost on HMI side - @5%s@'; 4098 'Maximum number of connections exceeded - @5%s@'; 4099 'Out of resources on PLC - @5%s@'; 4100 'Legitimation failed, invalid or missing password - @5%s@'; 4101 'Open request failed - @5%s@'; 4102 'Cannot connect to PLC - @5%s@'; 4103 'Open request could not be sent'; 4104 'root certificate expired for - @5%s@'; 4105 'PLC certificate untrusted for - @5%s@'

text list "SystemTextList_AllenBradleyDF1AlarmTextListCollection_9": 4096 'Connections: Connection to the PLC @5%s@ is lost'; 4097 'Connections: Connection to the HMI device @5%s@ is lost'; 4098 'Connections: Maximum number of connections exceeded - @5%s@'; 4099 'Out of resources on PLC - @5%s@'; 4100 'Legitimation failed, invalid or missing password - @5%s@'; 4101 'Request to open the connection failed - @5%s@'; 4102 'Connections: Cannot connect to PLC - @5%s@'; 4103 'Request to open the connection could not be sent'; 4104 'General certificate error for PLC - @5%s@'; 4105 'PLC certificate expired for PLC - @5%s@'; 4106 'PLC certificate is revoked for PLC - @5%s@'; 4107 'PLC certificate is untrustworthy. Manual trust is possible for - @5%s@'; 4108 'PLC certificate is untrustworthy. Manual trust is not possible for - @5%s@'

text list "SystemTextList_OmronEIPAlarmTextListCollection_6": 4096 'Connection lost on PLC side - @5%s@'; 4097 'Connection lost on HMI side - @5%s@'; 4098 'Maximum number of connections exceeded - @5%s@'; 4099 'Out of resources on PLC - @5%s@'; 4100 'Legitimation failed, invalid or missing password - @5%s@'; 4101 'Open request failed - @5%s@'; 4102 'Cannot connect to PLC - @5%s@'; 4103 'Open request could not be sent'; 4104 'root certificate expired for - @5%s@'; 4105 'PLC certificate untrusted for - @5%s@'

text list "SystemTextList_StdModbusTCPAlarmTextListCollection_5": 4096 'Connections: Connection to the PLC @5%s@ is lost'; 4097 'Connections: Connection to the HMI device @5%s@ is lost'; 4098 'Connections: Maximum number of connections exceeded - @5%s@'; 4099 'Out of resources on PLC - @5%s@'; 4100 'Legitimation failed, invalid or missing password - @5%s@'; 4101 'Request to open the connection failed - @5%s@'; 4102 'Connections: Cannot connect to PLC - @5%s@'; 4103 'Request to open the connection could not be sent'; 4104 'General certificate error for PLC - @5%s@'; 4105 'PLC certificate expired for PLC - @5%s@'; 4106 'PLC certificate is revoked for PLC - @5%s@'; 4107 'PLC certificate is untrustworthy. Manual trust is possible for - @5%s@'; 4108 'PLC certificate is untrustworthy. Manual trust is not possible for - @5%s@'

text list "SystemTextList_MitsubishiMCAlarmTextListCollection_4": 4096 'Connection lost on PLC side - @5%s@'; 4097 'Connection lost on HMI side - @5%s@'; 4098 'Maximum number of connections exceeded - @5%s@'; 4099 'Out of resources on PLC - @5%s@'; 4100 'Legitimation failed, invalid or missing password - @5%s@'; 4101 'Open request failed - @5%s@'; 4102 'Cannot connect to PLC - @5%s@'; 4103 'Open request could not be sent'; 4104 'root certificate expired for - @5%s@'; 4105 'PLC certificate untrusted for - @5%s@'

text list "SystemTextList_MitsubishiiQAlarmTextListCollection_3": 4096 'Connection lost on PLC side - @5%s@'; 4097 'Connection lost on HMI side - @5%s@'; 4098 'Maximum number of connections exceeded - @5%s@'; 4099 'Out of resources on PLC - @5%s@'; 4100 'Legitimation failed, invalid or missing password - @5%s@'; 4101 'Open request failed - @5%s@'; 4102 'Cannot connect to PLC - @5%s@'; 4103 'Open request could not be sent'; 4104 'root certificate expired for - @5%s@'; 4105 'PLC certificate untrusted for - @5%s@'

text list "SystemTextList_StdModbusRTUAlarmTextListCollection_8": 4096 'Connections: Connection to the PLC @5%s@ is lost'; 4097 'Connections: Connection to the HMI device @5%s@ is lost'; 4098 'Connections: Maximum number of connections exceeded - @5%s@'; 4099 'Out of resources on PLC - @5%s@'; 4100 'Legitimation failed, invalid or missing password - @5%s@'; 4101 'Request to open the connection failed - @5%s@'; 4102 'Connections: Cannot connect to PLC - @5%s@'; 4103 'Request to open the connection could not be sent'; 4104 'General certificate error for PLC - @5%s@'; 4105 'PLC certificate expired for PLC - @5%s@'; 4106 'PLC certificate is revoked for PLC - @5%s@'; 4107 'PLC certificate is untrustworthy. Manual trust is possible for - @5%s@'; 4108 'PLC certificate is untrustworthy. Manual trust is not possible for - @5%s@'

text list "SystemTextList_LogoAlarmTextListCollection_10": 4096 'Connections: Connection to the PLC @5%s@ is lost'; 4097 'Connections: Connection to the HMI device @5%s@ is lost'; 4098 'Connections: Maximum number of connections exceeded - @5%s@'; 4099 'Out of resources on PLC - @5%s@'; 4100 'Legitimation failed, invalid or missing password - @5%s@'; 4101 'Request to open the connection failed - @5%s@'; 4102 'Connections: Cannot connect to PLC - @5%s@'; 4103 'Request to open the connection could not be sent'; 4104 'General certificate error for PLC - @5%s@'; 4105 'PLC certificate expired for PLC - @5%s@'; 4106 'PLC certificate is revoked for PLC - @5%s@'; 4107 'PLC certificate is untrustworthy. Manual trust is possible for - @5%s@'; 4108 'PLC certificate is untrustworthy. Manual trust is not possible for - @5%s@'
*)